TYPE "Sensor U Shape Struct"
VERSION : 0.1


  STRUCT
   RISING_PULSE_1 : BOOL ;
   RISING_PULSE_2 : BOOL ;
   RISING_PULSE_3 : BOOL ;
   RISING_PULSE_4 : BOOL ;
   RISING_PULSE_5 : BOOL ;
   RISING_PULSE_6 : BOOL ;
   RISING_PULSE_7 : BOOL ;
   RISING_PULSE_8 : BOOL ;
   EVT_ACTIVE_0 : BOOL ;
   EVT_VALIDATED_0 : BOOL ;
   EVT_REJECTED_0 : BOOL ;
   EVT_ACTIVE_1 : BOOL ;
   BYPASS_LONG_0 : BOOL ;
   INIT_DONE : BOOL ;
   SPARE_1 : BOOL ;
   SPARE_2 : BOOL ;
   TMR_0_mS : INT ;
   TMR_1_mS : INT ;
   RESULT_SHORT_0 : INT ;
   VALIDATE_0_mS : INT ;
   DEBOUNCE_1_mS : INT ;
   COUNT_LIMIT : INT ;
  END_STRUCT ;
END_TYPE

